FUNCTION_BLOCK AlPgnRxNew_TP (* Receive a PGN of any length (also via transport protocol) into a byte array *)
  (* Standard: 61499-2; Description: Copyright (c) 2026 HR Agrartechnik GmbH This program and the accompanying materials are made available under the terms of the Eclipse Public License 2.0 which is available at https://www.eclipse.org/legal/epl-2.0/ SPDX-License-Identifier: EPL-2.0 Counterpart of AlPgnTxNew_TP. Data is an in/out byte array, e.g. from PROVIDE_ARR; its size limits the data that is kept. u16DaSize is the received length (up to 1785 bytes with TP, up to 65535 bytes with ETP). If it is larger than Data, the data is cut and OVERFLOW is TRUE. *)
  (* Version 1.0, 2026-11-13, Franz Höpfinger, HR Agrartechnik GmbH, Initial Version *)
  PACKAGE isobus::pgn::rx;
  IMPORT isobus::pgn::ISONETEVENT_T;
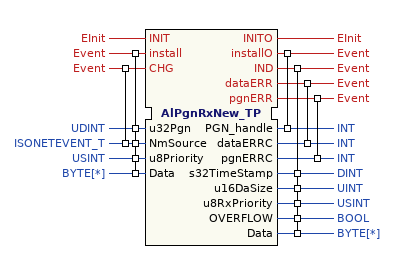
  EVENT_INPUT
    INIT : EInit; (* Service Initialization *)
    install WITH u32Pgn, NmSource, u8Priority, Data; (* installs a Receive PGN (RX) *)
    CHG WITH NmSource; (* Change source to NmSource.s16Handle *)
  END_EVENT
  EVENT_OUTPUT
    INITO : EInit; (* Initialization Confirm *)
    installO WITH PGN_handle; (* install Done *)
    IND WITH s32TimeStamp, u16DaSize, u8RxPriority, OVERFLOW, Data; (* Data was received *)
    dataERR WITH dataERRC;
    pgnERR WITH pgnERRC;
  END_EVENT
  VAR_INPUT
    u32Pgn : UDINT; (* PGN - Range: 0 - 0x3FFFF *)
    NmSource : isobus::pgn::ISONETEVENT_T; (* Define the Communication Partner *)
    u8Priority : USINT := 7; (* Priority given to the stack (0..7), not used as receive filter; received priority see u8RxPriority *)
  END_VAR
  VAR_OUTPUT
    PGN_handle : INT; (* PGN-handle on success, HANDLE_UNVALID in case of an error *)
    dataERRC : INT; (* dataERR error Code *)
    pgnERRC : INT; (* pgnERR error Code *)
    s32TimeStamp : DINT := -1; (* Time stamp of the message in ms *)
    u16DaSize : UINT; (* Received data length in bytes (0..65535) *)
    u8RxPriority : USINT; (* Priority of the received PGN *)
    OVERFLOW : BOOL; (* TRUE if more bytes were received than Data holds (Data is cut) *)
  END_VAR
  VAR_IN_OUT
    Data : ARRAY [*] OF BYTE; (* receive buffer, e.g. from PROVIDE_ARR *)
  END_VAR
END_FUNCTION_BLOCK
